// TIA Portal V19 export
DATA_BLOCK "RUA_R15_DB"   // DB56
// stored: InstanceOfName RUA_R15, InstanceOfType FB
"RUA_R15"
   // VAR
   //    START_Instance { S7_SetPoint := 'True'} : "START";
   //    "HEAT/COOL_Instance" { S7_SetPoint := 'True'} : "HEAT/COOL";
   //    "AUTO_COOLING_UTIITY SELECTION_Instance" { S7_SetPoint := 'True'} : "AUTO_COOLING_UTIITY SELECTION";
   //    AUTO_HEATING_SELECTION_Instance { S7_SetPoint := 'True'} : "AUTO_HEATING_SELECTION";
   //    COOLING_PROCESS_Instance { S7_SetPoint := 'True'} : "COOLING_PROCESS";
   //    HEATING_PROCEES_Instance { S7_SetPoint := 'True'} : "HEATING_PROCEES";
   //    RAMP_Instance { S7_SetPoint := 'True'} : "RAMP";
   //    "SEMI/_AUTO_Instance" { S7_SetPoint := 'True'} : "SEMI/_AUTO";
   // END_VAR
BEGIN
END_DATA_BLOCK
